Staubli VAL3: HWcheck.pgx

public program HWcheck()
  local num l_nNum
  local num l_nState
  local num l_nState1
  local string l_sState
begin
  //  rs:nHWState=$getState()
  //  l_nState=rs:nHWState
  //  if l_nState<0
  //    if !bReset
  //      l_nState=abs(l_nState)-90
  //      l_nState1=roundDown(l_nState)
  //      switch l_nState1
  //        case 0

  //          call rs:setAlarm(400,0)
  //        break
  //        case 1
  //          l_nNum= aioGet(ainRSI)
  //          if l_nNum!=0
  //            call rs:setAlarm(401,0)
  //          endIf
  //        break
  //        case 2
  //          call rs:setAlarm(402,0)
  //        break
  //        case 3
  //          call rs:setAlarm(403,0)
  //        break
  //        case 4
  //          call rs:setAlarm(404,0)
  //        break
  //        case 5
  //          call rs:setAlarm(405,0)
  //        break

  //      endSwitch
  //      bReset=true
  //    endIf
  //  else
  //    bReset=false
  //  endIf
end
